// TIA Portal V20 export
// export: Created 2026-10-12T05:42:34.286661Z, ExportSetting WithDefaults, DisplayName Totally Integrated Automation Portal, DisplayVersion V20, DisplayName TIA Portal Openness, DisplayVersion V20, DisplayName TIA Portal Teamcenter Gateway, DisplayVersion V20, DisplayName TIA Portal Version Control Interface, DisplayVersion V20, DisplayName SINAMICS Startdrive Advanced, DisplayVersion V20 SP1 Update 2, DisplayName SINAMICS Startdrive G110M, G120, G120C, G120D, G120P, G115D, DisplayVersion V20 SP1 Update 2, DisplayName SINAMICS Startdrive G130, G150, S120, S150, SINAMICS MV, G220, S200, S210, DisplayVersion V20 SP1 Update 2, DisplayName STEP 7 Professional, DisplayVersion V20, DisplayName STEP 7 Safety, DisplayVersion V20, DisplayName WinCC Basic/Comfort/Advanced, DisplayVersion V20, DisplayName WinCC Professional, DisplayVersion V20, DisplayName WinCC Unified, DisplayVersion V20
FUNCTION "F_PressDemoAwaitCycle" : Bool   // FC160, SCL
{ S7_Optimized_Access := 'TRUE' }
VERSION : 0.1
// stored: AutoNumber true, IsIECCheckEnabled false, SetENOAutomatically false, UDAEnableTagReadback false
   VAR_INPUT
      PartPresent : Bool;
      PartQuality : Bool;
      AirPressureOk : Bool;
      RequireTwoHandStart : Bool;
   END_VAR
   VAR_IN_OUT
      Seq : "FRK_SequenceCtx";
      Cycle : "ST_PressDemoCycle";
      Core : "FRK_Core";
      Unit : "FRK_Unit";
      Status : "ST_ModuleStatus";
      Part : "ST_PartContext";
      AlarmLog : "FRK_AlarmLog";
   END_VAR
   VAR_TEMP
      PartReady : Bool;
      AirReady : Bool;
      StartReady : Bool;
      Received : Bool;
   END_VAR
BEGIN

   #F_PressDemoAwaitCycle := FALSE;
   #Cycle.CycleCompleted := FALSE;
   IF #Unit.StopReq THEN
       "FRK_Complete"(Core := #Core,
                      Status := #Status);
       "FRK_SeqComplete"(Seq := #Seq);
       RETURN;
   END_IF;
   #PartReady := "FRK_SeqAwait"(Seq := #Seq, Label := 'project.condition.partPresent', Ok := #PartPresent AND #PartQuality);
   #AirReady := "FRK_SeqAwait"(Seq := #Seq, Label := 'project.condition.airPressureOk', Ok := #AirPressureOk);
   #StartReady := "FRK_SeqAwait"(Seq := #Seq, Label := 'project.condition.twoHandStart', Ok := #Seq.StartLatched OR NOT #RequireTwoHandStart);
   IF NOT (#PartReady AND #AirReady AND #StartReady) THEN
       RETURN;
   END_IF;
   IF NOT #Cycle.PartInMachine THEN
       #Received := "FRK_PartReceived"(Core := #Core, Unit := #Unit, Status := #Status, Part := #Part, AlarmLog := #AlarmLog);
       IF #Core.Exec = 3 THEN
           #Seq.Error := TRUE;
           #Seq.ErrorDiagnostic := #Status.Diagnostic;
           RETURN;
       END_IF;
       #Cycle.PartInMachine := TRUE;
   END_IF;
   #F_PressDemoAwaitCycle := TRUE;
END_FUNCTION
